// TIA Portal V21 export
Screen "T04_BtnSet"  1024x768, Number=24
  ScreenLayer 
    Button "P_Btn" at 0,0 size 100x30  TextOff="BTN", TextOn="BTN"
      EventHandler   EventType=Press
        FunctionCall "SetBit"
          FunctionParameter "Tag"  Tag=BtnStart
